Fanuc KAREL source: KA00145.KL

PROGRAM KA00145
%NOLOCKGROUP
VAR
  SRC: ARRAY[4] OF INTEGER
  DST: ARRAY[4] OF INTEGER
BEGIN
  DST = SRC
END KA00145
